(* PLC project Vn_leaf_assign, Beckhoff Automation GmbH TwinCAT PLC Control 3.5.13.21 *)
(* stored: creationDateTime 1970-01-01T00:00:00 *)

PROGRAM Vn_leaf_assign

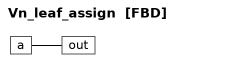
(* FBD diagram, written out as Structured Text *)
out := a;
END_PROGRAM
